(* IEC 61131-3 sources: llm-plc-st-eval/data/definitivo/gemini-3.1-pro-preview/I4/few_shot, 3 files *)

(* ---- ejec_1.st ---- *)
FUNCTION_BLOCK FB_EstrellaTriangulo
VAR_INPUT
    btnMarcha : BOOL; (* Boton de arranque *)
    btnParo : BOOL; (* Boton de parada *)
END_VAR
VAR_OUTPUT
    kM : BOOL; (* Contactor principal *)
    kY : BOOL; (* Contactor de estrella *)
    kD : BOOL; (* Contactor de triangulo *)
END_VAR
VAR
    enMarcha : BOOL; (* Memoria del estado del motor *)
    tEstrella : TON; (* Temporizador para la fase de estrella *)
    tMuerto : TON; (* Temporizador para el tiempo muerto *)
END_VAR

(* Control de marcha con prioridad a la parada *)
enMarcha := (btnMarcha OR enMarcha) AND NOT btnParo;

(* Temporizadores de transicion *)
tEstrella(IN := enMarcha, PT := T#8S);
tMuerto(IN := tEstrella.Q, PT := T#100MS);

(* Asignacion de salidas con enclavamiento de seguridad *)
kM := enMarcha;
kY := enMarcha AND NOT tEstrella.Q AND NOT kD;
kD := enMarcha AND tMuerto.Q AND NOT kY;
END_FUNCTION_BLOCK

(* ---- ejec_2.st ---- *)
FUNCTION_BLOCK FB_EstrellaTriangulo
VAR_INPUT
    btnMarcha : BOOL; (* Boton de arranque *)
    btnParo : BOOL;   (* Boton de parada *)
END_VAR
VAR_OUTPUT
    kM : BOOL; (* Contactor principal *)
    kY : BOOL; (* Contactor de estrella *)
    kD : BOOL; (* Contactor de triangulo *)
END_VAR
VAR
    enMarcha : BOOL; (* Memoria del estado de marcha *)
    tEstrella : TON; (* Temporizador de la fase estrella *)
    tMuerto : TON;   (* Temporizador del tiempo muerto *)
END_VAR

(* Control de marcha con prioridad a la parada *)
enMarcha := (enMarcha OR btnMarcha) AND NOT btnParo;

(* Temporizadores para la transicion *)
tEstrella(IN := enMarcha, PT := T#8S);
tMuerto(IN := tEstrella.Q, PT := T#100MS);

(* Activacion de contactores con enclavamiento mutuo de seguridad *)
kM := enMarcha;
kY := enMarcha AND NOT tEstrella.Q AND NOT kD;
kD := enMarcha AND tMuerto.Q AND NOT kY;
END_FUNCTION_BLOCK

(* ---- ejec_3.st ---- *)
FUNCTION_BLOCK FB_EstrellaTriangulo
VAR_INPUT
    btnMarcha : BOOL; (* Boton de arranque *)
    btnParo : BOOL;   (* Boton de parada *)
END_VAR
VAR_OUTPUT
    kM : BOOL; (* Contactor principal *)
    kY : BOOL; (* Contactor de estrella *)
    kD : BOOL; (* Contactor de triangulo *)
END_VAR
VAR
    tEstrella : TON; (* Temporizador de la fase estrella *)
    tMuerto : TON;   (* Temporizador del tiempo muerto *)
END_VAR

(* Memoria del contactor principal: se activa con marcha, se apaga con paro *)
kM := (btnMarcha OR kM) AND NOT btnParo;

(* Temporizadores para la transicion *)
tEstrella(IN := kM, PT := T#8S);
tMuerto(IN := tEstrella.Q, PT := T#100MS);

(* Contactor estrella: activo al inicio, se apaga a los 8s, interbloqueado con kD *)
kY := kM AND NOT tEstrella.Q AND NOT kD;

(* Contactor triangulo: activo tras el tiempo muerto, interbloqueado con kY *)
kD := kM AND tMuerto.Q AND NOT kY;
END_FUNCTION_BLOCK
